// TIA Portal V20 export
// export: Created 2026-11-08T12:00:00.0000000Z, ExportSetting None, DisplayName Totally Integrated Automation Portal, DisplayVersion V20, DisplayName STEP 7 Professional, DisplayVersion V20
FUNCTION_BLOCK "FB_Motor_DirectStart_LAD"   // FB20, LAD
TITLE = FB_Motor_DirectStart_LAD
{ S7_Optimized_Access := 'TRUE' }
// 电机直接起动带自锁与热过载保护（纯LAD实现）
// stored: AutoNumber false, MemoryReserve 10, SetENOAutomatically false
   VAR_INPUT
      startBtn : Bool;
      stopBtn : Bool;
      overloadNC : Bool;
   END_VAR
   VAR_OUTPUT
      motor : Bool;
   END_VAR
   VAR
      statMotor : Bool;
   END_VAR
BEGIN

REGION Network 1: 起保停自锁控制
   // 网络1：起保停自锁控制与停止/热过载保护
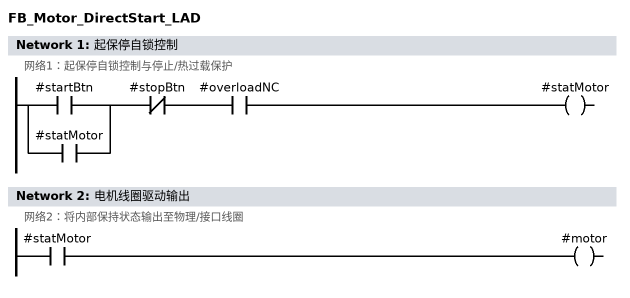
   RUNG wire#powerrail
      Contact( #startBtn )
      wire#w1
      I_Contact( #stopBtn )
      Contact( #overloadNC )
      Coil( #statMotor )
   END_RUNG
   RUNG wire#powerrail
      Contact( #statMotor )
   END_RUNG wire#w1
   // the same network as SCL:
   #statMotor := (#startBtn OR #statMotor) AND NOT #stopBtn AND #overloadNC;
END_REGION

REGION Network 2: 电机线圈驱动输出
   // 网络2：将内部保持状态输出至物理/接口线圈
   RUNG wire#powerrail
      Contact( #statMotor )
      Coil( #motor )
   END_RUNG
   // the same network as SCL:
   #motor := #statMotor;
END_REGION
END_FUNCTION_BLOCK
